FUNCTION_BLOCK clear_err
VAR_INPUT
END_VAR
VAR_OUTPUT
END_VAR
VAR
	i:INT;
	step:INT:=0;
	settle_timer:TON;
	all_powered:BOOL;
	has_err:BOOL;
END_VAR

(* 
Post-error recovery:
  - keep the handle input frozen
  - cold start or a fresh _init cycle must return to _init until self-check is completed
  - otherwise wait until errors are gone and all axes are powered again
  - then reinitialize handle references from the current position
*)

has_err := FALSE;
FOR i:=1 TO 7 DO
	IF G.axis[i].Status.Error OR G.power_output[i].Error OR G.reset_output[i].Error THEN
		has_err := TRUE;
		EXIT;
	END_IF
END_FOR

all_powered := TRUE;
FOR i:=1 TO 7 DO
	IF NOT G.power_output[i].Done THEN
		all_powered := FALSE;
		EXIT;
	END_IF
END_FOR

G.estop_hold_req := TRUE;

CASE step OF
0:
	FOR i:=1 TO 7 DO
		G.SetPointGenEnable[i].Execute := FALSE;
		G.SetPointGenDisable[i].Execute := FALSE;
		G.axis_Reset[i].Execute := FALSE;
	END_FOR
	settle_timer(IN:=FALSE);
	step := 1;

1:
	IF has_err THEN
		settle_timer(IN:=FALSE);
		step := 0;
		G.gen_state := _err;
		RETURN;
	END_IF

	IF NOT G.self_check_done THEN
		settle_timer(IN:=FALSE);
		step := 0;
		G.gen_state := _init;
		RETURN;
	END_IF

	IF NOT all_powered THEN
		FOR i:=1 TO 7 DO
			G.power_[i].Enable := TRUE;
		END_FOR
		settle_timer(IN:=FALSE);
		RETURN;
	END_IF

	settle_timer(IN:=TRUE, PT:=T#200MS);
	IF settle_timer.Q THEN
		settle_timer(IN:=FALSE);
		step := 0;
		G.handle_reinit_req := TRUE;
		G.gen_state := _handle;
	END_IF
END_CASE

END_FUNCTION_BLOCK

(* stored: Version 1.1.0.1, ProductVersion 3.1.4024.15
   POU clear_err: Id {b44b79d2-0ec3-452a-abc9-d2df60552efa}, SpecialFunc None *)
